(* PLC project Plc, Beckhoff Automation GmbH TwinCAT PLC Control 3.5.21.61 *)
(* stored: creationDateTime 2026-10-21T14:48:56.5320043, modificationDateTime 2026-10-21T14:48:56.5369587 *)

INTERFACE I_Module
// Runs one cycle; FALSE while in error
METHOD Execute : BOOL
VAR_INPUT
	eCmd : E_Command;
END_VAR
END_METHOD
// N175 retest marker
METHOD GetStatus : ST_ModuleStatus
END_METHOD
END_INTERFACE
